KUKA KRL program: pick_place.src, pick_place.dat

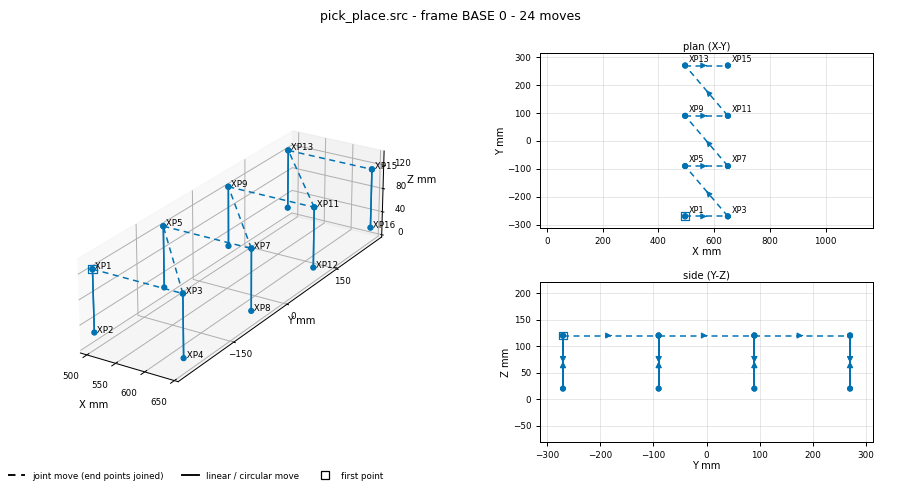
[picture p0: tool path of pick_place.src in frame BASE 0, 24 of 26 moves have a stored position in this frame; points joined in program order, loops and branches not executed]
--- pick_place.src ---
&ACCESS RVP
&REL 1
&PARAM EDITMASK = *
&PARAM TEMPLATE = C:\KRC\Roboter\Template\vorgabe
&PARAM DISKPATH = KRC:\R1\Program
DEF pick_place( )
; KR 6 R900 sixx (AGILUS) 픽 앤 플레이스 예제 (RobotEmulator 자동 생성)
; 그리퍼: Robotiq 2F-85 Adaptive
; $OUT[1]=그리퍼 닫기, $OUT[2]=그리퍼 열기, $IN[1]=닫힘 확인, $IN[2]=열림 확인
  ;FOLD INI;%{PE}
    ;FOLD BASISTECH INI
      GLOBAL INTERRUPT DECL 3 WHEN $STOPMESS==TRUE DO IR_STOPM ( )
      INTERRUPT ON 3
      BAS (#INITMOV,0 )
    ;ENDFOLD (BASISTECH INI)
    ;FOLD USER INI
      ;Make your modifications here
      nPart = 0
    ;ENDFOLD (USER INI)
  ;ENDFOLD (INI)

  ;FOLD PTP HOME  Vel= 100 % DEFAULT;%{PE}%MKUKATPBASIS,%CMOVE,%VPTP,%P 1:PTP, 2:HOME, 3:, 5:100, 7:DEFAULT
  $BWDSTART = FALSE
  PDAT_ACT=PDEFAULT
  FDAT_ACT=FHOME
  BAS (#PTP_PARAMS,100 )
  $H_POS=XHOME
  PTP  XHOME
  ;ENDFOLD
  GripOpen()

  ; ---- 공작물 W1 (1/4) ----
  ;FOLD PTP P1 Vel=100 % PDAT1 Tool[1]:gripper Base[0];%{PE}%R 8.3.48,%MKUKATPBASIS,%CMOVE,%VPTP,%P 1:PTP, 2:P1, 3:, 5:100, 7:PDAT1
  $BWDSTART=FALSE
  PDAT_ACT=PPDAT1
  FDAT_ACT=FP1
  BAS(#PTP_PARAMS,100)
  PTP XP1
  ;ENDFOLD
  ;FOLD LIN P2 Vel=0.3 m/s CPDAT1 Tool[1]:gripper Base[0];%{PE}%R 8.3.48,%MKUKATPBASIS,%CMOVE,%VLIN,%P 1:LIN, 2:P2, 3:, 5:0.3, 7:CPDAT1
  $BWDSTART=FALSE
  LDAT_ACT=LCPDAT1
  FDAT_ACT=FP2
  BAS(#CP_PARAMS,0.3)
  LIN XP2
  ;ENDFOLD
  GripClose()
  ;FOLD LIN P1 Vel=0.5 m/s CPDAT2 Tool[1]:gripper Base[0];%{PE}%R 8.3.48,%MKUKATPBASIS,%CMOVE,%VLIN,%P 1:LIN, 2:P1, 3:, 5:0.5, 7:CPDAT2
  $BWDSTART=FALSE
  LDAT_ACT=LCPDAT2
  FDAT_ACT=FP1
  BAS(#CP_PARAMS,0.5)
  LIN XP1
  ;ENDFOLD
  ;FOLD PTP P3 Vel=100 % PDAT2 Tool[1]:gripper Base[0];%{PE}%R 8.3.48,%MKUKATPBASIS,%CMOVE,%VPTP,%P 1:PTP, 2:P3, 3:, 5:100, 7:PDAT2
  $BWDSTART=FALSE
  PDAT_ACT=PPDAT2
  FDAT_ACT=FP3
  BAS(#PTP_PARAMS,100)
  PTP XP3
  ;ENDFOLD
  ;FOLD LIN P4 Vel=0.3 m/s CPDAT3 Tool[1]:gripper Base[0];%{PE}%R 8.3.48,%MKUKATPBASIS,%CMOVE,%VLIN,%P 1:LIN, 2:P4, 3:, 5:0.3, 7:CPDAT3
  $BWDSTART=FALSE
  LDAT_ACT=LCPDAT3
  FDAT_ACT=FP4
  BAS(#CP_PARAMS,0.3)
  LIN XP4
  ;ENDFOLD
  GripOpen()
  ;FOLD LIN P3 Vel=0.5 m/s CPDAT4 Tool[1]:gripper Base[0];%{PE}%R 8.3.48,%MKUKATPBASIS,%CMOVE,%VLIN,%P 1:LIN, 2:P3, 3:, 5:0.5, 7:CPDAT4
  $BWDSTART=FALSE
  LDAT_ACT=LCPDAT4
  FDAT_ACT=FP3
  BAS(#CP_PARAMS,0.5)
  LIN XP3
  ;ENDFOLD
  nPart = nPart + 1

  ; ---- 공작물 W2 (2/4) ----
  ;FOLD PTP P5 Vel=100 % PDAT3 Tool[1]:gripper Base[0];%{PE}%R 8.3.48,%MKUKATPBASIS,%CMOVE,%VPTP,%P 1:PTP, 2:P5, 3:, 5:100, 7:PDAT3
  $BWDSTART=FALSE
  PDAT_ACT=PPDAT3
  FDAT_ACT=FP5
  BAS(#PTP_PARAMS,100)
  PTP XP5
  ;ENDFOLD
  ;FOLD LIN P6 Vel=0.3 m/s CPDAT5 Tool[1]:gripper Base[0];%{PE}%R 8.3.48,%MKUKATPBASIS,%CMOVE,%VLIN,%P 1:LIN, 2:P6, 3:, 5:0.3, 7:CPDAT5
  $BWDSTART=FALSE
  LDAT_ACT=LCPDAT5
  FDAT_ACT=FP6
  BAS(#CP_PARAMS,0.3)
  LIN XP6
  ;ENDFOLD
  GripClose()
  ;FOLD LIN P5 Vel=0.5 m/s CPDAT6 Tool[1]:gripper Base[0];%{PE}%R 8.3.48,%MKUKATPBASIS,%CMOVE,%VLIN,%P 1:LIN, 2:P5, 3:, 5:0.5, 7:CPDAT6
  $BWDSTART=FALSE
  LDAT_ACT=LCPDAT6
  FDAT_ACT=FP5
  BAS(#CP_PARAMS,0.5)
  LIN XP5
  ;ENDFOLD
  ;FOLD PTP P7 Vel=100 % PDAT4 Tool[1]:gripper Base[0];%{PE}%R 8.3.48,%MKUKATPBASIS,%CMOVE,%VPTP,%P 1:PTP, 2:P7, 3:, 5:100, 7:PDAT4
  $BWDSTART=FALSE
  PDAT_ACT=PPDAT4
  FDAT_ACT=FP7
  BAS(#PTP_PARAMS,100)
  PTP XP7
  ;ENDFOLD
  ;FOLD LIN P8 Vel=0.3 m/s CPDAT7 Tool[1]:gripper Base[0];%{PE}%R 8.3.48,%MKUKATPBASIS,%CMOVE,%VLIN,%P 1:LIN, 2:P8, 3:, 5:0.3, 7:CPDAT7
  $BWDSTART=FALSE
  LDAT_ACT=LCPDAT7
  FDAT_ACT=FP8
  BAS(#CP_PARAMS,0.3)
  LIN XP8
  ;ENDFOLD
  GripOpen()
  ;FOLD LIN P7 Vel=0.5 m/s CPDAT8 Tool[1]:gripper Base[0];%{PE}%R 8.3.48,%MKUKATPBASIS,%CMOVE,%VLIN,%P 1:LIN, 2:P7, 3:, 5:0.5, 7:CPDAT8
  $BWDSTART=FALSE
  LDAT_ACT=LCPDAT8
  FDAT_ACT=FP7
  BAS(#CP_PARAMS,0.5)
  LIN XP7
  ;ENDFOLD
  nPart = nPart + 1

  ; ---- 공작물 W3 (3/4) ----
  ;FOLD PTP P9 Vel=100 % PDAT5 Tool[1]:gripper Base[0];%{PE}%R 8.3.48,%MKUKATPBASIS,%CMOVE,%VPTP,%P 1:PTP, 2:P9, 3:, 5:100, 7:PDAT5
  $BWDSTART=FALSE
  PDAT_ACT=PPDAT5
  FDAT_ACT=FP9
  BAS(#PTP_PARAMS,100)
  PTP XP9
  ;ENDFOLD
  ;FOLD LIN P10 Vel=0.3 m/s CPDAT9 Tool[1]:gripper Base[0];%{PE}%R 8.3.48,%MKUKATPBASIS,%CMOVE,%VLIN,%P 1:LIN, 2:P10, 3:, 5:0.3, 7:CPDAT9
  $BWDSTART=FALSE
  LDAT_ACT=LCPDAT9
  FDAT_ACT=FP10
  BAS(#CP_PARAMS,0.3)
  LIN XP10
  ;ENDFOLD
  GripClose()
  ;FOLD LIN P9 Vel=0.5 m/s CPDAT10 Tool[1]:gripper Base[0];%{PE}%R 8.3.48,%MKUKATPBASIS,%CMOVE,%VLIN,%P 1:LIN, 2:P9, 3:, 5:0.5, 7:CPDAT10
  $BWDSTART=FALSE
  LDAT_ACT=LCPDAT10
  FDAT_ACT=FP9
  BAS(#CP_PARAMS,0.5)
  LIN XP9
  ;ENDFOLD
  ;FOLD PTP P11 Vel=100 % PDAT6 Tool[1]:gripper Base[0];%{PE}%R 8.3.48,%MKUKATPBASIS,%CMOVE,%VPTP,%P 1:PTP, 2:P11, 3:, 5:100, 7:PDAT6
  $BWDSTART=FALSE
  PDAT_ACT=PPDAT6
  FDAT_ACT=FP11
  BAS(#PTP_PARAMS,100)
  PTP XP11
  ;ENDFOLD
  ;FOLD LIN P12 Vel=0.3 m/s CPDAT11 Tool[1]:gripper Base[0];%{PE}%R 8.3.48,%MKUKATPBASIS,%CMOVE,%VLIN,%P 1:LIN, 2:P12, 3:, 5:0.3, 7:CPDAT11
  $BWDSTART=FALSE
  LDAT_ACT=LCPDAT11
  FDAT_ACT=FP12
  BAS(#CP_PARAMS,0.3)
  LIN XP12
  ;ENDFOLD
  GripOpen()
  ;FOLD LIN P11 Vel=0.5 m/s CPDAT12 Tool[1]:gripper Base[0];%{PE}%R 8.3.48,%MKUKATPBASIS,%CMOVE,%VLIN,%P 1:LIN, 2:P11, 3:, 5:0.5, 7:CPDAT12
  $BWDSTART=FALSE
  LDAT_ACT=LCPDAT12
  FDAT_ACT=FP11
  BAS(#CP_PARAMS,0.5)
  LIN XP11
  ;ENDFOLD
  nPart = nPart + 1

  ; ---- 공작물 W4 (4/4) ----
  ;FOLD PTP P13 Vel=100 % PDAT7 Tool[1]:gripper Base[0];%{PE}%R 8.3.48,%MKUKATPBASIS,%CMOVE,%VPTP,%P 1:PTP, 2:P13, 3:, 5:100, 7:PDAT7
  $BWDSTART=FALSE
  PDAT_ACT=PPDAT7
  FDAT_ACT=FP13
  BAS(#PTP_PARAMS,100)
  PTP XP13
  ;ENDFOLD
  ;FOLD LIN P14 Vel=0.3 m/s CPDAT13 Tool[1]:gripper Base[0];%{PE}%R 8.3.48,%MKUKATPBASIS,%CMOVE,%VLIN,%P 1:LIN, 2:P14, 3:, 5:0.3, 7:CPDAT13
  $BWDSTART=FALSE
  LDAT_ACT=LCPDAT13
  FDAT_ACT=FP14
  BAS(#CP_PARAMS,0.3)
  LIN XP14
  ;ENDFOLD
  GripClose()
  ;FOLD LIN P13 Vel=0.5 m/s CPDAT14 Tool[1]:gripper Base[0];%{PE}%R 8.3.48,%MKUKATPBASIS,%CMOVE,%VLIN,%P 1:LIN, 2:P13, 3:, 5:0.5, 7:CPDAT14
  $BWDSTART=FALSE
  LDAT_ACT=LCPDAT14
  FDAT_ACT=FP13
  BAS(#CP_PARAMS,0.5)
  LIN XP13
  ;ENDFOLD
  ;FOLD PTP P15 Vel=100 % PDAT8 Tool[1]:gripper Base[0];%{PE}%R 8.3.48,%MKUKATPBASIS,%CMOVE,%VPTP,%P 1:PTP, 2:P15, 3:, 5:100, 7:PDAT8
  $BWDSTART=FALSE
  PDAT_ACT=PPDAT8
  FDAT_ACT=FP15
  BAS(#PTP_PARAMS,100)
  PTP XP15
  ;ENDFOLD
  ;FOLD LIN P16 Vel=0.3 m/s CPDAT15 Tool[1]:gripper Base[0];%{PE}%R 8.3.48,%MKUKATPBASIS,%CMOVE,%VLIN,%P 1:LIN, 2:P16, 3:, 5:0.3, 7:CPDAT15
  $BWDSTART=FALSE
  LDAT_ACT=LCPDAT15
  FDAT_ACT=FP16
  BAS(#CP_PARAMS,0.3)
  LIN XP16
  ;ENDFOLD
  GripOpen()
  ;FOLD LIN P15 Vel=0.5 m/s CPDAT16 Tool[1]:gripper Base[0];%{PE}%R 8.3.48,%MKUKATPBASIS,%CMOVE,%VLIN,%P 1:LIN, 2:P15, 3:, 5:0.5, 7:CPDAT16
  $BWDSTART=FALSE
  LDAT_ACT=LCPDAT16
  FDAT_ACT=FP15
  BAS(#CP_PARAMS,0.5)
  LIN XP15
  ;ENDFOLD
  nPart = nPart + 1

  ;FOLD PTP HOME  Vel= 100 % DEFAULT;%{PE}%MKUKATPBASIS,%CMOVE,%VPTP,%P 1:PTP, 2:HOME, 3:, 5:100, 7:DEFAULT
  $BWDSTART = FALSE
  PDAT_ACT=PDEFAULT
  FDAT_ACT=FHOME
  BAS (#PTP_PARAMS,100 )
  $H_POS=XHOME
  PTP  XHOME
  ;ENDFOLD
  MsgNotify("픽 앤 플레이스 완료")
END

DEF GripClose( )
  ;FOLD OUT 2 'Gripper open' State=FALSE ;%{PE}%R 8.3.48,%MKUKATPBASIS,%COUT,%VOUTX,%P 2:2, 3:Gripper open, 5:FALSE, 6:
  $OUT[2]=FALSE
  ;ENDFOLD
  ;FOLD OUT 1 'Gripper close' State=TRUE ;%{PE}%R 8.3.48,%MKUKATPBASIS,%COUT,%VOUTX,%P 2:1, 3:Gripper close, 5:TRUE, 6:
  $OUT[1]=TRUE
  ;ENDFOLD
  ;FOLD WAIT FOR IN 1 'Gripper closed' ;%{PE}%R 8.3.48,%MKUKATPBASIS,%CEXT_WAIT_FOR,%VEXT_WAIT_FOR,%P 2:, 4:, 5:$IN, 6:1, 7:Gripper closed, 9:
  WAIT FOR  ( $IN[1] )
  ;ENDFOLD
  ;FOLD WAIT Time=0.2 sec;%{PE}%R 8.3.48,%MKUKATPBASIS,%CWAIT,%VWAIT,%P 2:0.2
  WAIT SEC 0.2
  ;ENDFOLD
END

DEF GripOpen( )
  ;FOLD OUT 1 'Gripper close' State=FALSE ;%{PE}%R 8.3.48,%MKUKATPBASIS,%COUT,%VOUTX,%P 2:1, 3:Gripper close, 5:FALSE, 6:
  $OUT[1]=FALSE
  ;ENDFOLD
  ;FOLD OUT 2 'Gripper open' State=TRUE ;%{PE}%R 8.3.48,%MKUKATPBASIS,%COUT,%VOUTX,%P 2:2, 3:Gripper open, 5:TRUE, 6:
  $OUT[2]=TRUE
  ;ENDFOLD
  ;FOLD WAIT FOR IN 2 'Gripper opened' ;%{PE}%R 8.3.48,%MKUKATPBASIS,%CEXT_WAIT_FOR,%VEXT_WAIT_FOR,%P 2:, 4:, 5:$IN, 6:2, 7:Gripper opened, 9:
  WAIT FOR  ( $IN[2] )
  ;ENDFOLD
  $OUT[2]=FALSE
  WAIT SEC 0.2
END

--- pick_place.dat ---
&ACCESS RVP
&REL 1
&PARAM EDITMASK = *
&PARAM TEMPLATE = C:\KRC\Roboter\Template\vorgabe
&PARAM DISKPATH = KRC:\R1\Program
DEFDAT  pick_place
;FOLD EXTERNAL DECLARATIONS;%{PE}%MKUKATPBASIS,%CEXT,%VCOMMON,%P
;FOLD BASISTECH EXT;%{PE}%MKUKATPBASIS,%CEXT,%VEXT,%P
EXT  BAS (BAS_COMMAND  :IN,REAL  :IN )
DECL INT SUCCESS
;ENDFOLD (BASISTECH EXT)
;FOLD USER EXT;%{E}%MKUKATPUSER,%CEXT,%VEXT,%P
;Make your modifications here
DECL INT nPart=0
;ENDFOLD (USER EXT)
;ENDFOLD (EXTERNAL DECLARATIONS)
DECL E6POS XP1={X 495.825,Y -270.45,Z 120.0,A 180.000,B 0.0,C 180.000,S 2,T 2,E1 0.0,E2 0.0,E3 0.0,E4 0.0,E5 0.0,E6 0.0}
DECL FDAT FP1={TOOL_NO 1,BASE_NO 0,IPO_FRAME #BASE,POINT2[] " "}
DECL E6POS XP2={X 495.825,Y -270.45,Z 20.0,A 180.000,B 0.0,C 180.000,S 2,T 2,E1 0.0,E2 0.0,E3 0.0,E4 0.0,E5 0.0,E6 0.0}
DECL FDAT FP2={TOOL_NO 1,BASE_NO 0,IPO_FRAME #BASE,POINT2[] " "}
DECL E6POS XP3={X 649.08,Y -270.45,Z 120.0,A 180.000,B 0.0,C 180.000,S 2,T 2,E1 0.0,E2 0.0,E3 0.0,E4 0.0,E5 0.0,E6 0.0}
DECL FDAT FP3={TOOL_NO 1,BASE_NO 0,IPO_FRAME #BASE,POINT2[] " "}
DECL E6POS XP4={X 649.08,Y -270.45,Z 20.0,A 180.000,B 0.0,C 180.000,S 2,T 2,E1 0.0,E2 0.0,E3 0.0,E4 0.0,E5 0.0,E6 0.0}
DECL FDAT FP4={TOOL_NO 1,BASE_NO 0,IPO_FRAME #BASE,POINT2[] " "}
DECL E6POS XP5={X 495.825,Y -90.15,Z 120.0,A 180.000,B 0.0,C 180.000,S 2,T 2,E1 0.0,E2 0.0,E3 0.0,E4 0.0,E5 0.0,E6 0.0}
DECL FDAT FP5={TOOL_NO 1,BASE_NO 0,IPO_FRAME #BASE,POINT2[] " "}
DECL E6POS XP6={X 495.825,Y -90.15,Z 20.0,A 180.000,B 0.0,C 180.000,S 2,T 2,E1 0.0,E2 0.0,E3 0.0,E4 0.0,E5 0.0,E6 0.0}
DECL FDAT FP6={TOOL_NO 1,BASE_NO 0,IPO_FRAME #BASE,POINT2[] " "}
DECL E6POS XP7={X 649.08,Y -90.15,Z 120.0,A 180.000,B 0.0,C 180.000,S 2,T 2,E1 0.0,E2 0.0,E3 0.0,E4 0.0,E5 0.0,E6 0.0}
DECL FDAT FP7={TOOL_NO 1,BASE_NO 0,IPO_FRAME #BASE,POINT2[] " "}
DECL E6POS XP8={X 649.08,Y -90.15,Z 20.0,A 180.000,B 0.0,C 180.000,S 2,T 2,E1 0.0,E2 0.0,E3 0.0,E4 0.0,E5 0.0,E6 0.0}
DECL FDAT FP8={TOOL_NO 1,BASE_NO 0,IPO_FRAME #BASE,POINT2[] " "}
DECL E6POS XP9={X 495.825,Y 90.15,Z 120.0,A 180.000,B 0.0,C 180.000,S 2,T 35,E1 0.0,E2 0.0,E3 0.0,E4 0.0,E5 0.0,E6 0.0}
DECL FDAT FP9={TOOL_NO 1,BASE_NO 0,IPO_FRAME #BASE,POINT2[] " "}
DECL E6POS XP10={X 495.825,Y 90.15,Z 20.0,A 180.000,B 0.0,C 180.000,S 2,T 35,E1 0.0,E2 0.0,E3 0.0,E4 0.0,E5 0.0,E6 0.0}
DECL FDAT FP10={TOOL_NO 1,BASE_NO 0,IPO_FRAME #BASE,POINT2[] " "}
DECL E6POS XP11={X 649.08,Y 90.15,Z 120.0,A 180.000,B 0.0,C 180.000,S 2,T 35,E1 0.0,E2 0.0,E3 0.0,E4 0.0,E5 0.0,E6 0.0}
DECL FDAT FP11={TOOL_NO 1,BASE_NO 0,IPO_FRAME #BASE,POINT2[] " "}
DECL E6POS XP12={X 649.08,Y 90.15,Z 20.0,A 180.000,B 0.0,C 180.000,S 2,T 35,E1 0.0,E2 0.0,E3 0.0,E4 0.0,E5 0.0,E6 0.0}
DECL FDAT FP12={TOOL_NO 1,BASE_NO 0,IPO_FRAME #BASE,POINT2[] " "}
DECL E6POS XP13={X 495.825,Y 270.45,Z 120.0,A 180.000,B 0.0,C 180.000,S 2,T 35,E1 0.0,E2 0.0,E3 0.0,E4 0.0,E5 0.0,E6 0.0}
DECL FDAT FP13={TOOL_NO 1,BASE_NO 0,IPO_FRAME #BASE,POINT2[] " "}
DECL E6POS XP14={X 495.825,Y 270.45,Z 20.0,A 180.000,B 0.0,C 180.000,S 2,T 35,E1 0.0,E2 0.0,E3 0.0,E4 0.0,E5 0.0,E6 0.0}
DECL FDAT FP14={TOOL_NO 1,BASE_NO 0,IPO_FRAME #BASE,POINT2[] " "}
DECL E6POS XP15={X 649.08,Y 270.45,Z 120.0,A 180.000,B 0.0,C 180.000,S 2,T 35,E1 0.0,E2 0.0,E3 0.0,E4 0.0,E5 0.0,E6 0.0}
DECL FDAT FP15={TOOL_NO 1,BASE_NO 0,IPO_FRAME #BASE,POINT2[] " "}
DECL E6POS XP16={X 649.08,Y 270.45,Z 20.0,A 180.000,B 0.0,C 180.000,S 2,T 35,E1 0.0,E2 0.0,E3 0.0,E4 0.0,E5 0.0,E6 0.0}
DECL FDAT FP16={TOOL_NO 1,BASE_NO 0,IPO_FRAME #BASE,POINT2[] " "}
DECL PDAT PPDAT1={VEL 100.000,ACC 100.000,APO_DIST 100.000,APO_MODE #CDIS,GEAR_JERK 50.0000,EXAX_IGN 0}
DECL LDAT LCPDAT1={VEL 0.3,ACC 100.000,APO_DIST 100.000,APO_FAC 50.0000,AXIS_VEL 100.000,AXIS_ACC 100.000,ORI_TYP #VAR,CIRC_TYP #BASE,JERK_FAC 50.0000,GEAR_JERK 50.0000,EXAX_IGN 0}
DECL LDAT LCPDAT2={VEL 0.5,ACC 100.000,APO_DIST 100.000,APO_FAC 50.0000,AXIS_VEL 100.000,AXIS_ACC 100.000,ORI_TYP #VAR,CIRC_TYP #BASE,JERK_FAC 50.0000,GEAR_JERK 50.0000,EXAX_IGN 0}
DECL PDAT PPDAT2={VEL 100.000,ACC 100.000,APO_DIST 100.000,APO_MODE #CDIS,GEAR_JERK 50.0000,EXAX_IGN 0}
DECL LDAT LCPDAT3={VEL 0.3,ACC 100.000,APO_DIST 100.000,APO_FAC 50.0000,AXIS_VEL 100.000,AXIS_ACC 100.000,ORI_TYP #VAR,CIRC_TYP #BASE,JERK_FAC 50.0000,GEAR_JERK 50.0000,EXAX_IGN 0}
DECL LDAT LCPDAT4={VEL 0.5,ACC 100.000,APO_DIST 100.000,APO_FAC 50.0000,AXIS_VEL 100.000,AXIS_ACC 100.000,ORI_TYP #VAR,CIRC_TYP #BASE,JERK_FAC 50.0000,GEAR_JERK 50.0000,EXAX_IGN 0}
DECL PDAT PPDAT3={VEL 100.000,ACC 100.000,APO_DIST 100.000,APO_MODE #CDIS,GEAR_JERK 50.0000,EXAX_IGN 0}
DECL LDAT LCPDAT5={VEL 0.3,ACC 100.000,APO_DIST 100.000,APO_FAC 50.0000,AXIS_VEL 100.000,AXIS_ACC 100.000,ORI_TYP #VAR,CIRC_TYP #BASE,JERK_FAC 50.0000,GEAR_JERK 50.0000,EXAX_IGN 0}
DECL LDAT LCPDAT6={VEL 0.5,ACC 100.000,APO_DIST 100.000,APO_FAC 50.0000,AXIS_VEL 100.000,AXIS_ACC 100.000,ORI_TYP #VAR,CIRC_TYP #BASE,JERK_FAC 50.0000,GEAR_JERK 50.0000,EXAX_IGN 0}
DECL PDAT PPDAT4={VEL 100.000,ACC 100.000,APO_DIST 100.000,APO_MODE #CDIS,GEAR_JERK 50.0000,EXAX_IGN 0}
DECL LDAT LCPDAT7={VEL 0.3,ACC 100.000,APO_DIST 100.000,APO_FAC 50.0000,AXIS_VEL 100.000,AXIS_ACC 100.000,ORI_TYP #VAR,CIRC_TYP #BASE,JERK_FAC 50.0000,GEAR_JERK 50.0000,EXAX_IGN 0}
DECL LDAT LCPDAT8={VEL 0.5,ACC 100.000,APO_DIST 100.000,APO_FAC 50.0000,AXIS_VEL 100.000,AXIS_ACC 100.000,ORI_TYP #VAR,CIRC_TYP #BASE,JERK_FAC 50.0000,GEAR_JERK 50.0000,EXAX_IGN 0}
DECL PDAT PPDAT5={VEL 100.000,ACC 100.000,APO_DIST 100.000,APO_MODE #CDIS,GEAR_JERK 50.0000,EXAX_IGN 0}
DECL LDAT LCPDAT9={VEL 0.3,ACC 100.000,APO_DIST 100.000,APO_FAC 50.0000,AXIS_VEL 100.000,AXIS_ACC 100.000,ORI_TYP #VAR,CIRC_TYP #BASE,JERK_FAC 50.0000,GEAR_JERK 50.0000,EXAX_IGN 0}
DECL LDAT LCPDAT10={VEL 0.5,ACC 100.000,APO_DIST 100.000,APO_FAC 50.0000,AXIS_VEL 100.000,AXIS_ACC 100.000,ORI_TYP #VAR,CIRC_TYP #BASE,JERK_FAC 50.0000,GEAR_JERK 50.0000,EXAX_IGN 0}
DECL PDAT PPDAT6={VEL 100.000,ACC 100.000,APO_DIST 100.000,APO_MODE #CDIS,GEAR_JERK 50.0000,EXAX_IGN 0}
DECL LDAT LCPDAT11={VEL 0.3,ACC 100.000,APO_DIST 100.000,APO_FAC 50.0000,AXIS_VEL 100.000,AXIS_ACC 100.000,ORI_TYP #VAR,CIRC_TYP #BASE,JERK_FAC 50.0000,GEAR_JERK 50.0000,EXAX_IGN 0}
DECL LDAT LCPDAT12={VEL 0.5,ACC 100.000,APO_DIST 100.000,APO_FAC 50.0000,AXIS_VEL 100.000,AXIS_ACC 100.000,ORI_TYP #VAR,CIRC_TYP #BASE,JERK_FAC 50.0000,GEAR_JERK 50.0000,EXAX_IGN 0}
DECL PDAT PPDAT7={VEL 100.000,ACC 100.000,APO_DIST 100.000,APO_MODE #CDIS,GEAR_JERK 50.0000,EXAX_IGN 0}
DECL LDAT LCPDAT13={VEL 0.3,ACC 100.000,APO_DIST 100.000,APO_FAC 50.0000,AXIS_VEL 100.000,AXIS_ACC 100.000,ORI_TYP #VAR,CIRC_TYP #BASE,JERK_FAC 50.0000,GEAR_JERK 50.0000,EXAX_IGN 0}
DECL LDAT LCPDAT14={VEL 0.5,ACC 100.000,APO_DIST 100.000,APO_FAC 50.0000,AXIS_VEL 100.000,AXIS_ACC 100.000,ORI_TYP #VAR,CIRC_TYP #BASE,JERK_FAC 50.0000,GEAR_JERK 50.0000,EXAX_IGN 0}
DECL PDAT PPDAT8={VEL 100.000,ACC 100.000,APO_DIST 100.000,APO_MODE #CDIS,GEAR_JERK 50.0000,EXAX_IGN 0}
DECL LDAT LCPDAT15={VEL 0.3,ACC 100.000,APO_DIST 100.000,APO_FAC 50.0000,AXIS_VEL 100.000,AXIS_ACC 100.000,ORI_TYP #VAR,CIRC_TYP #BASE,JERK_FAC 50.0000,GEAR_JERK 50.0000,EXAX_IGN 0}
DECL LDAT LCPDAT16={VEL 0.5,ACC 100.000,APO_DIST 100.000,APO_FAC 50.0000,AXIS_VEL 100.000,AXIS_ACC 100.000,ORI_TYP #VAR,CIRC_TYP #BASE,JERK_FAC 50.0000,GEAR_JERK 50.0000,EXAX_IGN 0}
ENDDAT
